// TIA Portal V20 export
TYPE "Störmeldung_PN"
   STRUCT
      Störmeldung_PN : Array[0..127] of Bool;
   END_STRUCT;
END_TYPE
